FUNCTION_BLOCK ABSTRACT FB_SafetyBase EXTENDS KOSTAL_AF2024_Core_Station.FB_Station_Free IMPLEMENTS I_Safety
VAR
	_inHold				: BOOL;
	_isSafe				: BOOL;
	_doorLock			: BOOL;
	_isDoorUsed			: BOOL:= TRUE;
	_isDoorSafe			: BOOL;
	_manual				: BOOL;
	_tempIsSafe			: BOOL;
	_logMessageStart	: BOOL;
	(* Hmi *)
	_Hmi_station		: KOSTAL_AF2024_HMI_WinHMI.FB_Page_Station;
	_E_Text				: T_E_text_Safety;
END_VAR

METHOD PROTECTED ABSTRACT  _handleSafety 
VAR_INPUT
END_VAR
END_METHOD

METHOD PROTECTED _hmiDefine
VAR_INPUT
END_VAR
_Hmi_station.Name:= _Name;

_Hmi_station.Text.line_01:= _condition.Message.line_01;
_Hmi_station.Text.line_02:= _condition.Message.line_02;
_Hmi_station.Text.line_03:= _condition.Message.line_03;

_Hmi_station.Button_Escape.Visible:= (_condition.isError() OR _Hmi_station.Button_Escape.Sign) AND _manual;
_Hmi_station.Button_Escape.Text:= _Text.GetText(Number:= _E_Text.reset);

_Hmi_station.Status.CopyFrom(IN:= _condition);

_Hmi_station.FBmain();
END_METHOD

METHOD PROTECTED _logStart
VAR_INPUT
END_VAR
IF _logMessageStart AND _Text.State.ready AND (_Text.LoadedLanguage <> '') THEN
	IF _log("===START===") THEN
		_logMessageStart:= FALSE;
	END_IF
	
	IF _tempIsSafe THEN 
		_log(Text:= _Text.GetText(Number:= _E_Text.safetyOk));
	ELSE
		_log(Text:= _Text.GetText(Number:= _E_Text.safetyNok));
	END_IF
END_IF
END_METHOD

METHOD PROTECTED _resetCondition 
VAR_INPUT
END_VAR
IF _condition.isError() THEN
	IF _Hmi_station.Button_Escape.Pulse THEN
		_condition.clear();
	END_IF
ELSE
	_condition.clear();
END_IF
END_METHOD

PROPERTY PUBLIC doorLock : BOOL
GET
doorLock:= _doorLock;
END_GET
SET
_doorLock:= doorLock;
END_SET
END_PROPERTY

METHOD FB_init : BOOL
VAR_INPUT
	bInitRetains : BOOL; // if TRUE, the retain variables are initialized (warm start / cold start)
	bInCopyCode : BOOL;  // if TRUE, the instance afterwards gets moved into the copy code (online change)
	ID_Name			: KOSTAL_AF2024_Core_Settings.T_MaxString;
	ID_Key			: DINT;
	CommonText		: KOSTAL_AF2024_Core_Text.I_Text;
	textPath		: KOSTAL_AF2024_Core_Settings.T_MaxString_UTF8;
END_VAR
_TextPath:= textPath;
END_METHOD

METHOD PUBLIC FBmain
VAR_INPUT
END_VAR
IF NOT _parameterControl() THEN RETURN; END_IF
 
_hmiDefine();

IF NOT _TextReader() THEN RETURN; END_IF;

_logStart();
_handleSafety();
_resetCondition();
_tempIsSafe:= NOT _condition.isError();

(* Log if safety state changed *)
IF _isSafe <> _tempIsSafe THEN
	IF _tempIsSafe THEN			
		_log(_Text.GetText(_E_text.safetyOk));
	ELSE							
		_log(_condition.Message.toString());				
	END_IF
END_IF

_isSafe:= _tempIsSafe;

IF _isSafe THEN	
	_message.clear();
	_message.line_01:= _Text.GetText(Number:= _E_text.safetyOk);
	_condition.setMessage(
		priority:= _condition.PriorityLevel_Info, 
		message	:= _message);
END_IF
END_METHOD

PROPERTY inHold : BOOL
GET
inHold:= _inHold;
END_GET
END_PROPERTY

PROPERTY isDoorSafe : BOOL
GET
isDoorSafe:= _isDoorSafe;
END_GET
END_PROPERTY

PROPERTY isDoorUsed : BOOL
GET
isDoorUsed:= _isDoorUsed;
END_GET
END_PROPERTY

PROPERTY isSafe : BOOL
GET
isSafe:= _isSafe;
END_GET
END_PROPERTY

PROPERTY PUBLIC manual : BOOL
GET
manual := _manual;
END_GET
SET
_manual:= manual;
END_SET
END_PROPERTY

END_FUNCTION_BLOCK

(* stored: Version 1.1.0.1, ProductVersion 3.1.4024.12
   POU FB_SafetyBase: Id {12bade05-da6f-4709-92e0-138c674938c3}, SpecialFunc None
   Folder Private: Id {88030c51-4729-4a31-8c0f-dd20f061485c}
   Folder Property: Id {191e8cbf-d21b-4a8a-ba34-ee36284c8b26}
   Method _handleSafety: Id {7df14ae7-5b1f-4cd5-b48f-db327fe3265c}
   Method _hmiDefine: Id {69d24df7-3eb4-424b-a243-8f202c54ed24}
   Method _logStart: Id {c42151e0-164b-412f-854c-fc50caf71b9d}
   Method _resetCondition: Id {dc02b2bc-ebda-4b19-986d-a81c01eaa0a1}
   Property doorLock: Id {13d368e7-a983-479d-8fd8-068a0b9cd829}
   Get Get: Id {c2cf3276-0dc2-4f67-a108-8d35332db5da}
   Set Set: Id {8a1e11fb-2f91-422e-992c-2d258eae0145}
   Method FB_init: Id {cce0d010-45e2-493d-bc29-dd2af3806d59}
   Method FBmain: Id {645b2cb8-bff5-46c3-a477-544e29134ee7}
   Property inHold: Id {065ef20f-1211-4cda-8bf0-49df9f2a4ee3}
   Get Get: Id {ef0b982d-eb5a-4b3c-98cf-51a6d9eedc91}
   Property isDoorSafe: Id {affcff9d-fdf9-401a-a228-18a0aa9f5bde}
   Get Get: Id {019d570a-26b2-4997-aaf6-e20e0b755092}
   Property isDoorUsed: Id {f4a7b5c6-afda-44ea-b144-5ddaf3f8d41e}
   Get Get: Id {00e5b138-8de1-4d6b-bd72-a7d652478473}
   Property isSafe: Id {3f10ae2f-4e65-4f5c-87a0-25babdfe5316}
   Get Get: Id {e29e2e6a-ff3d-4f43-a02d-ebc20e949737}
   Property manual: Id {75062206-38e6-47ac-bef8-a7289ba56dc5}
   Get Get: Id {3c2d1efa-d8d4-4ac6-8216-7dd081e0a000}
   Set Set: Id {67cb55cf-5fe0-477e-bafe-ea4c2c012881} *)
